(* IEC 61131-3 sources: trust-platform/examples/network_canvas_demo/src, 2 files *)

(* ---- config.st ---- *)
CONFIGURATION Config
VAR_GLOBAL
    conveyor_speed : REAL := 1.5;
    running : BOOL := FALSE;
    line_state : INT := 1;
END_VAR
RESOURCE CommRes ON PLC
    TASK MainTask (INTERVAL := T#10ms, PRIORITY := 1);
    PROGRAM Main WITH MainTask : Main;
END_RESOURCE
END_CONFIGURATION

(* ---- main.st ---- *)
PROGRAM Main
VAR_EXTERNAL
    conveyor_speed : REAL;
    running : BOOL;
    line_state : INT;
END_VAR

running := TRUE;
IF conveyor_speed < 2.0 THEN
    conveyor_speed := conveyor_speed + 0.1;
END_IF;
line_state := 1;
END_PROGRAM
